// SIMATIC S7-200 project (STEP 7-Micro/WIN), CPU 224XP CN REL 02.01

SYMBOL_TABLE USUARIO1
SO               I0.3     // Sensor de Objetos (Detecta la pieza para iniciar la seleccion)
S_I              I0.4     // Sensor de fibra Optica (clasificacion de materiales)
SM               I0.5     // Sensor magnetico (clasificacion de materiales)
S1               I0.7     // Sensor de retorno del cilindro 1
S2               I1.0     // Sensor de retorno del cilindro 2
S3               I1.1     // Sensor de retorno del cilindro 3
SBB1             I1.3     // Pulsador de Marcha
SBB2             I1.2     // Pulsador de Paro
QS               I1.4     // Zeta de emergencia
SA               I1.5     // Selector rotatorio
am               Q0.0     // Motor
C_1              Q0.4     // cilindro neumatico 1
C_2              Q0.5     // cilindro neumatico 2
C_3              Q0.6     // cilindro neumatico 3
HL1              Q0.7     // Lampara de señalizacion amarilla
HL2              Q1.0     // Lampara de señalizacion verde
HL3              Q1.1     // Lampara de señalizacion roja
E0               M0.0     // Estado 0
E1               M0.1     // Estado 1
E2               M0.2     // Estado 2
E3               M0.3     // Estado 3
E4               M0.4     // Estado 4
E5               M0.5     // Estado 5
E6               M0.6     // Estado 6
E7               M0.7     // Estado 7
E8               M1.0     // Estado 8
E9               M1.1     // Estado 9
E10              M1.2     // Estado 10
E11              M1.3     // Estado 11
E12              M1.4     // Estado 12
E13              M1.5     // Estado 13
E14              M1.6     // Estado 14
EM               M1.7     // Variable para paro momentaneo
MOTOR            M2.0     // Variable para activacion o desactivacion del motor
E15              M2.1     // Estado 15
E16              M2.2     // Estado 16
C_C0             VD110
C_C1             VD100
r_k              VD190
m_k              VD120
m_k_1            VD130
m_k_2            VD140
e_k              VD150
e_k_1            VD160
e_k_2            VD170
Ao               VD200
Bo               VD210
Co               VD220
Do               VD230
Eo               VD240
L_k              VD180
set_point        VD90
END_SYMBOL_TABLE

ORGANIZATION_BLOCK PRINCIPAL:OB1
TITLE=UNIDAD DE SELECCION
BEGIN
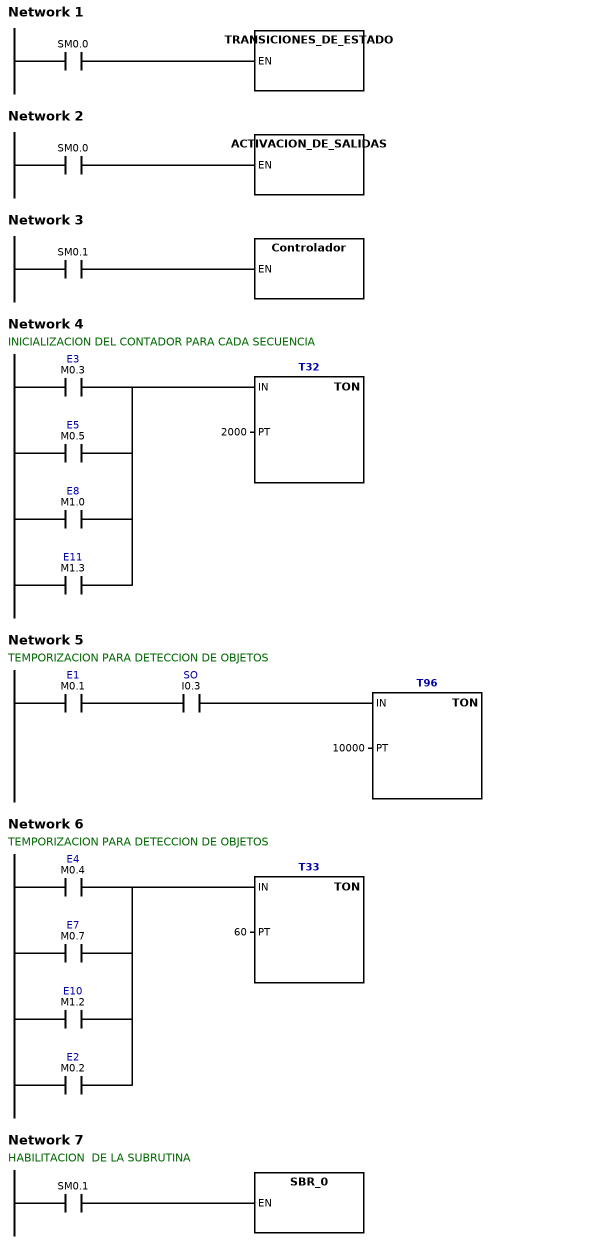
Network 1
LD     SM0.0
CALL   TRANSICIONES_DE_ESTADO:SBR1
Network 2
LD     SM0.0
CALL   ACTIVACION_DE_SALIDAS:SBR2
Network 3
LD     SM0.1
CALL   Controlador:SBR3
Network 4
// INICIALIZACION DEL CONTADOR PARA CADA SECUENCIA 
LD     E3:M0.3
O      E5:M0.5
O      E8:M1.0
O      E11:M1.3
TON    T32, 2000
Network 5
// TEMPORIZACION PARA DETECCION DE OBJETOS
LD     E1:M0.1
A      SO:I0.3
TON    T96, 10000
Network 6
// TEMPORIZACION PARA DETECCION DE OBJETOS
LD     E4:M0.4
O      E7:M0.7
O      E10:M1.2
O      E2:M0.2
TON    T33, 60
Network 7
// HABILITACION  DE LA SUBRUTINA
LD     SM0.1
CALL   SBR_0:SBR0
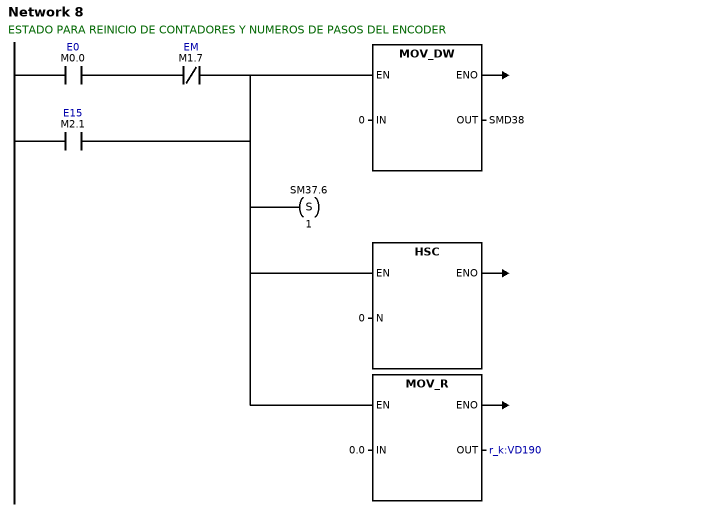
Network 8
// ESTADO PARA REINICIO DE CONTADORES Y NUMEROS DE PASOS DEL ENCODER
LD     E0:M0.0
AN     EM:M1.7
O      E15:M2.1
MOVD   0, SMD38
S      SM37.6, 1
HSC    0
MOVR   0.0, r_k:VD190
END_ORGANIZATION_BLOCK

SUBROUTINE_BLOCK SBR_0:SBR0
TITLE=COMENTARIOS DE LA SUBRUTINA
BEGIN
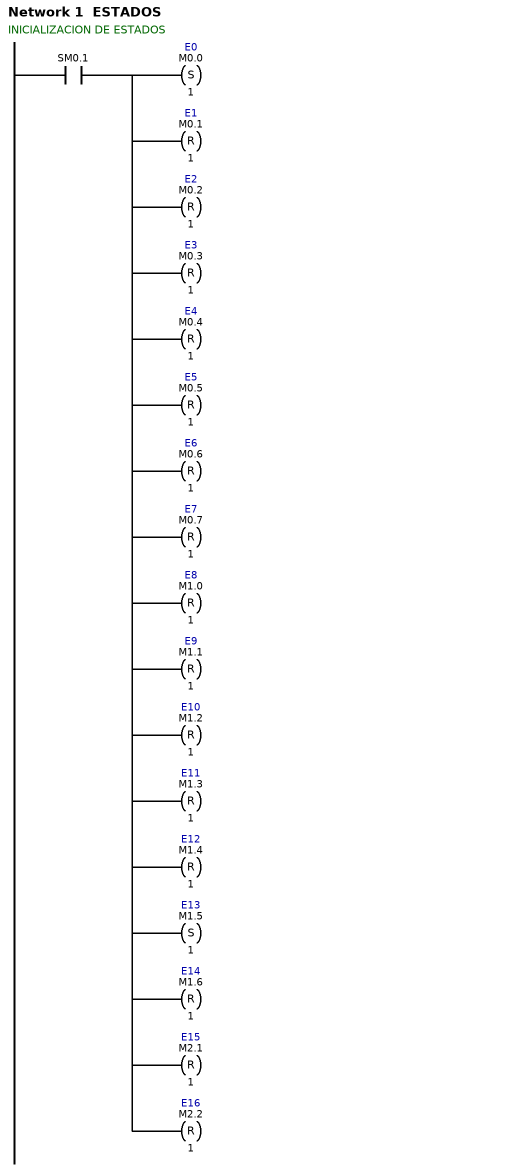
Network 1 // ESTADOS
// INICIALIZACION DE ESTADOS
LD     SM0.1
S      E0:M0.0, 1
R      E1:M0.1, 1
R      E2:M0.2, 1
R      E3:M0.3, 1
R      E4:M0.4, 1
R      E5:M0.5, 1
R      E6:M0.6, 1
R      E7:M0.7, 1
R      E8:M1.0, 1
R      E9:M1.1, 1
R      E10:M1.2, 1
R      E11:M1.3, 1
R      E12:M1.4, 1
S      E13:M1.5, 1
R      E14:M1.6, 1
R      E15:M2.1, 1
R      E16:M2.2, 1
END_SUBROUTINE_BLOCK

SUBROUTINE_BLOCK TRANSICIONES_DE_ESTADO:SBR1
TITLE=TRANSICIONES DE ESTADO
BEGIN
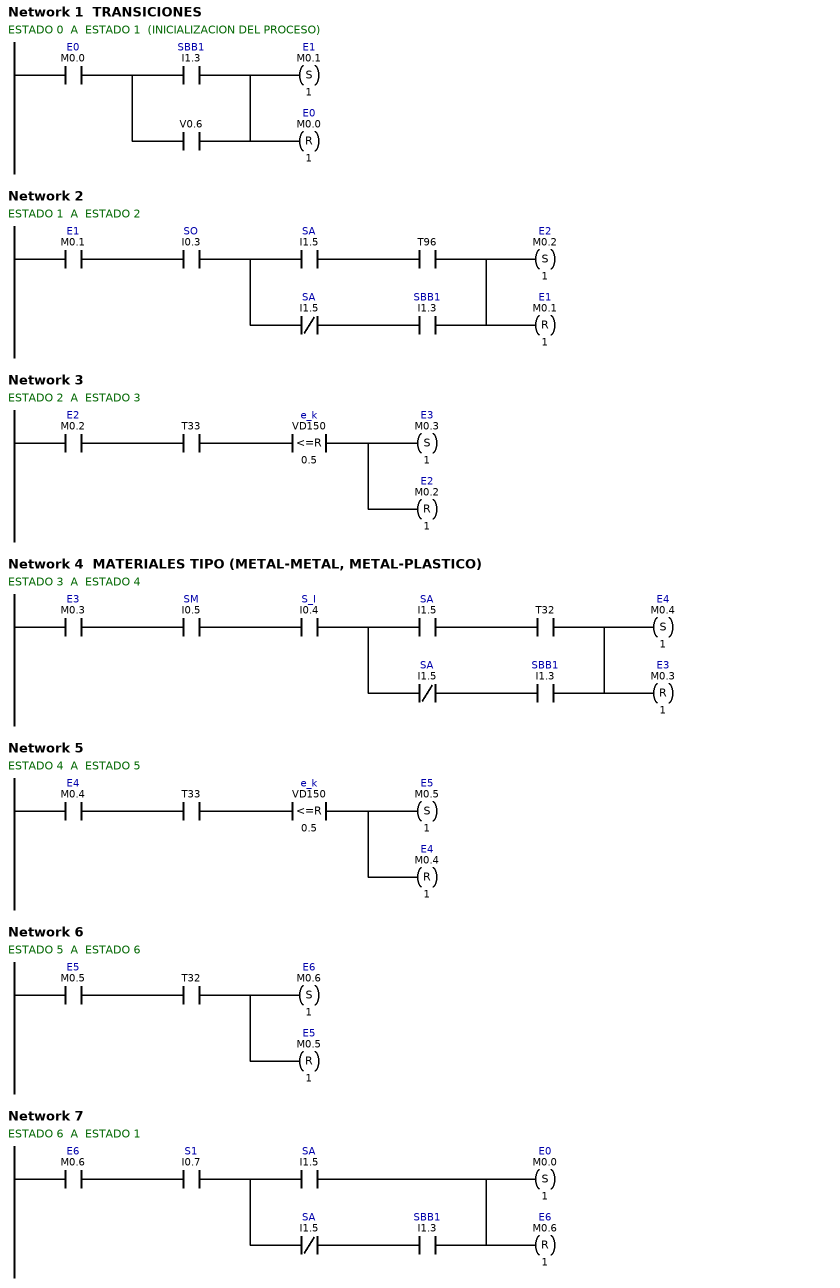
Network 1 // TRANSICIONES
// ESTADO 0  A  ESTADO 1  (INICIALIZACION DEL PROCESO)
LD     E0:M0.0
LD     SBB1:I1.3
O      V0.6
ALD
S      E1:M0.1, 1
R      E0:M0.0, 1
Network 2
// ESTADO 1  A  ESTADO 2 
LD     E1:M0.1
A      SO:I0.3
LD     SA:I1.5
A      T96
LDN    SA:I1.5
A      SBB1:I1.3
OLD
ALD
S      E2:M0.2, 1
R      E1:M0.1, 1
Network 3
// ESTADO 2  A  ESTADO 3
LD     E2:M0.2
A      T33
AR<=   e_k:VD150, 0.5
S      E3:M0.3, 1
R      E2:M0.2, 1
Network 4 // MATERIALES TIPO (METAL-METAL, METAL-PLASTICO)
// ESTADO 3  A  ESTADO 4
LD     E3:M0.3
A      SM:I0.5
A      S_I:I0.4
LD     SA:I1.5
A      T32
LDN    SA:I1.5
A      SBB1:I1.3
OLD
ALD
S      E4:M0.4, 1
R      E3:M0.3, 1
Network 5
// ESTADO 4  A  ESTADO 5
LD     E4:M0.4
A      T33
AR<=   e_k:VD150, 0.5
S      E5:M0.5, 1
R      E4:M0.4, 1
Network 6
// ESTADO 5  A  ESTADO 6
LD     E5:M0.5
A      T32
S      E6:M0.6, 1
R      E5:M0.5, 1
Network 7
// ESTADO 6  A  ESTADO 1
LD     E6:M0.6
A      S1:I0.7
LD     SA:I1.5
LDN    SA:I1.5
A      SBB1:I1.3
OLD
ALD
S      E0:M0.0, 1
R      E6:M0.6, 1
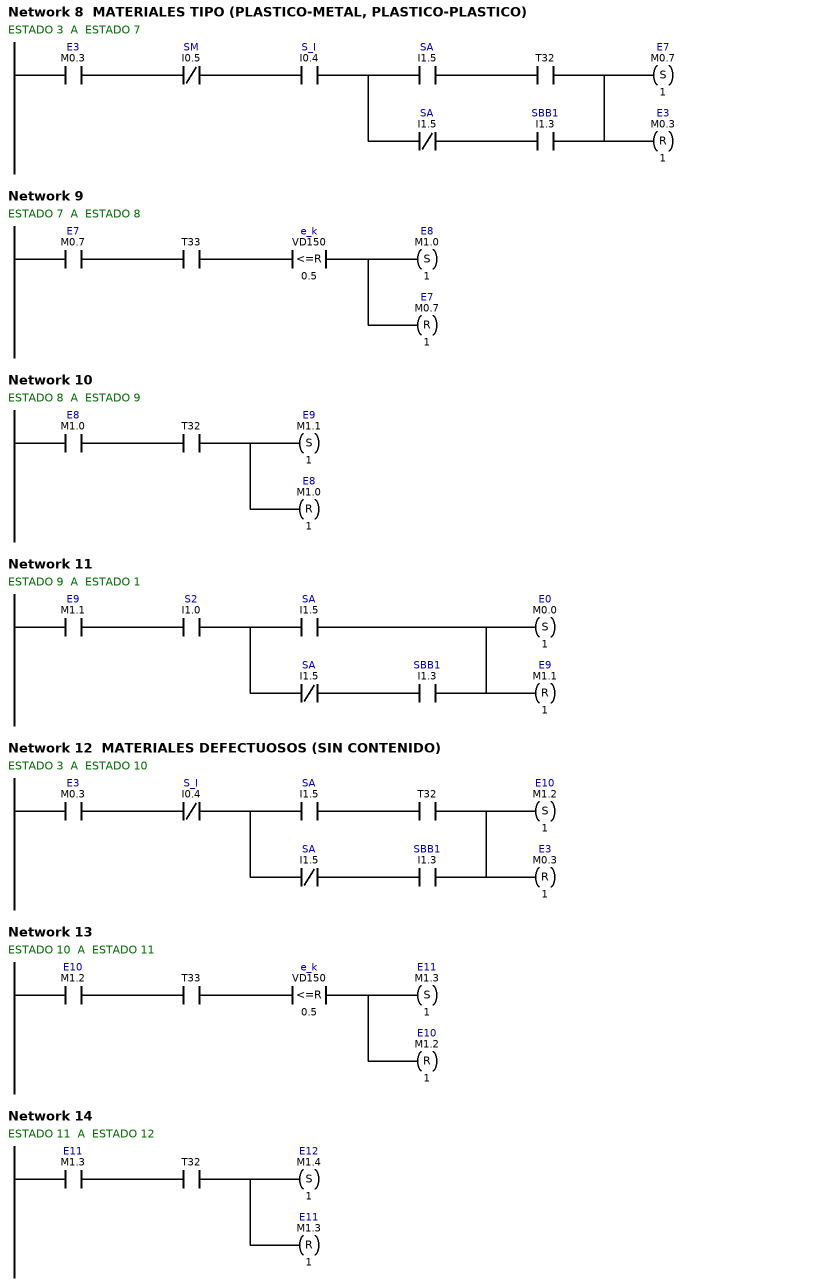
Network 8 // MATERIALES TIPO (PLASTICO-METAL, PLASTICO-PLASTICO)
// ESTADO 3  A  ESTADO 7
LD     E3:M0.3
AN     SM:I0.5
A      S_I:I0.4
LD     SA:I1.5
A      T32
LDN    SA:I1.5
A      SBB1:I1.3
OLD
ALD
S      E7:M0.7, 1
R      E3:M0.3, 1
Network 9
// ESTADO 7  A  ESTADO 8
LD     E7:M0.7
A      T33
AR<=   e_k:VD150, 0.5
S      E8:M1.0, 1
R      E7:M0.7, 1
Network 10
// ESTADO 8  A  ESTADO 9
LD     E8:M1.0
A      T32
S      E9:M1.1, 1
R      E8:M1.0, 1
Network 11
// ESTADO 9  A  ESTADO 1
LD     E9:M1.1
A      S2:I1.0
LD     SA:I1.5
LDN    SA:I1.5
A      SBB1:I1.3
OLD
ALD
S      E0:M0.0, 1
R      E9:M1.1, 1
Network 12 // MATERIALES DEFECTUOSOS (SIN CONTENIDO)
// ESTADO 3  A  ESTADO 10 
LD     E3:M0.3
AN     S_I:I0.4
LD     SA:I1.5
A      T32
LDN    SA:I1.5
A      SBB1:I1.3
OLD
ALD
S      E10:M1.2, 1
R      E3:M0.3, 1
Network 13
// ESTADO 10  A  ESTADO 11
LD     E10:M1.2
A      T33
AR<=   e_k:VD150, 0.5
S      E11:M1.3, 1
R      E10:M1.2, 1
Network 14
// ESTADO 11  A  ESTADO 12
LD     E11:M1.3
A      T32
S      E12:M1.4, 1
R      E11:M1.3, 1
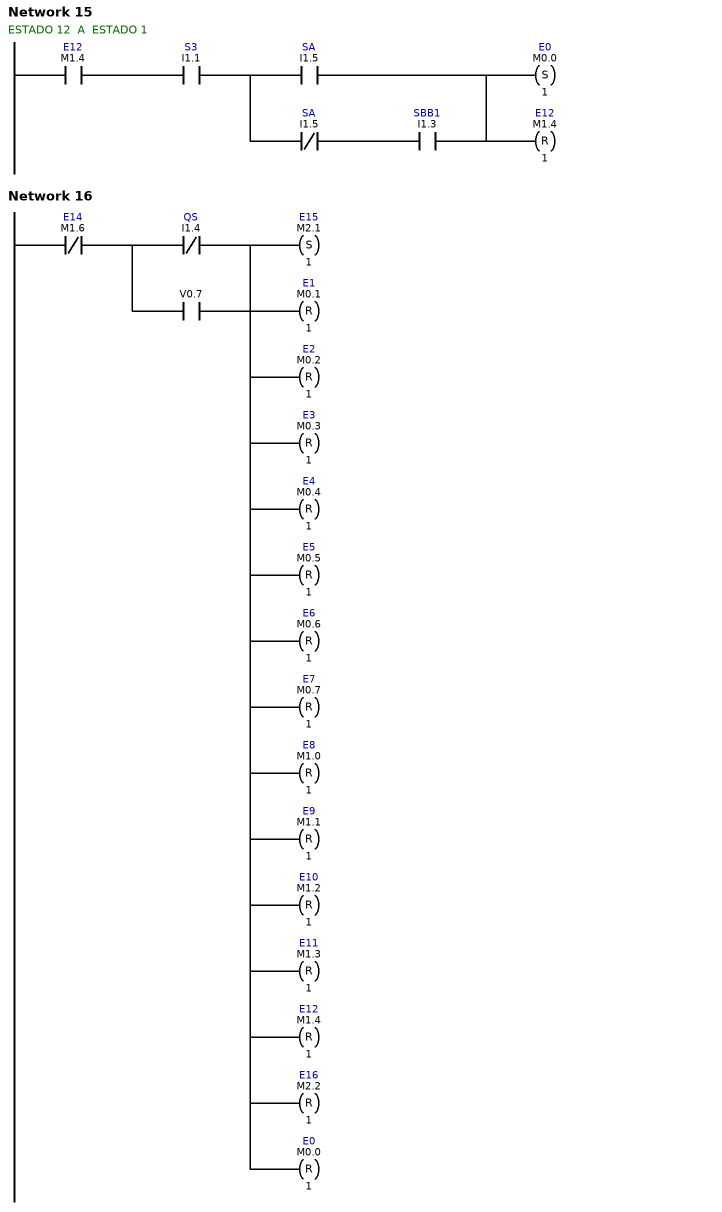
Network 15
// ESTADO 12  A  ESTADO 1
LD     E12:M1.4
A      S3:I1.1
LD     SA:I1.5
LDN    SA:I1.5
A      SBB1:I1.3
OLD
ALD
S      E0:M0.0, 1
R      E12:M1.4, 1
Network 16
LDN    E14:M1.6
LDN    QS:I1.4
O      V0.7
ALD
S      E15:M2.1, 1
R      E1:M0.1, 1
R      E2:M0.2, 1
R      E3:M0.3, 1
R      E4:M0.4, 1
R      E5:M0.5, 1
R      E6:M0.6, 1
R      E7:M0.7, 1
R      E8:M1.0, 1
R      E9:M1.1, 1
R      E10:M1.2, 1
R      E11:M1.3, 1
R      E12:M1.4, 1
R      E16:M2.2, 1
R      E0:M0.0, 1
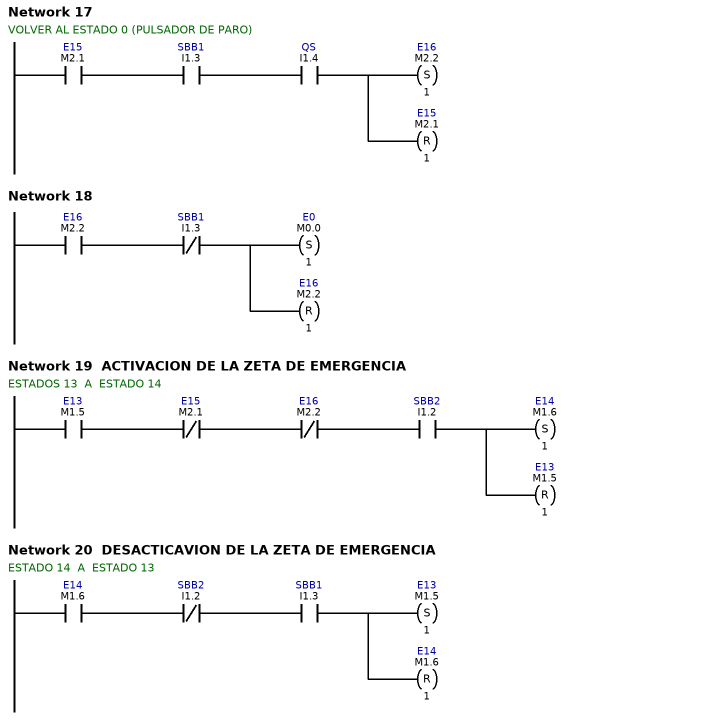
Network 17
// VOLVER AL ESTADO 0 (PULSADOR DE PARO)
LD     E15:M2.1
A      SBB1:I1.3
A      QS:I1.4
S      E16:M2.2, 1
R      E15:M2.1, 1
Network 18
LD     E16:M2.2
AN     SBB1:I1.3
S      E0:M0.0, 1
R      E16:M2.2, 1
Network 19 // ACTIVACION DE LA ZETA DE EMERGENCIA
// ESTADOS 13  A  ESTADO 14
LD     E13:M1.5
AN     E15:M2.1
AN     E16:M2.2
A      SBB2:I1.2
S      E14:M1.6, 1
R      E13:M1.5, 1
Network 20 // DESACTICAVION DE LA ZETA DE EMERGENCIA
// ESTADO 14  A  ESTADO 13
LD     E14:M1.6
AN     SBB2:I1.2
A      SBB1:I1.3
S      E13:M1.5, 1
R      E14:M1.6, 1
Network 21 // Título de segmento
// Comentario de segmento
END_SUBROUTINE_BLOCK

SUBROUTINE_BLOCK ACTIVACION_DE_SALIDAS:SBR2
TITLE=COMENTARIOS DE LA SUBRUTINA
BEGIN
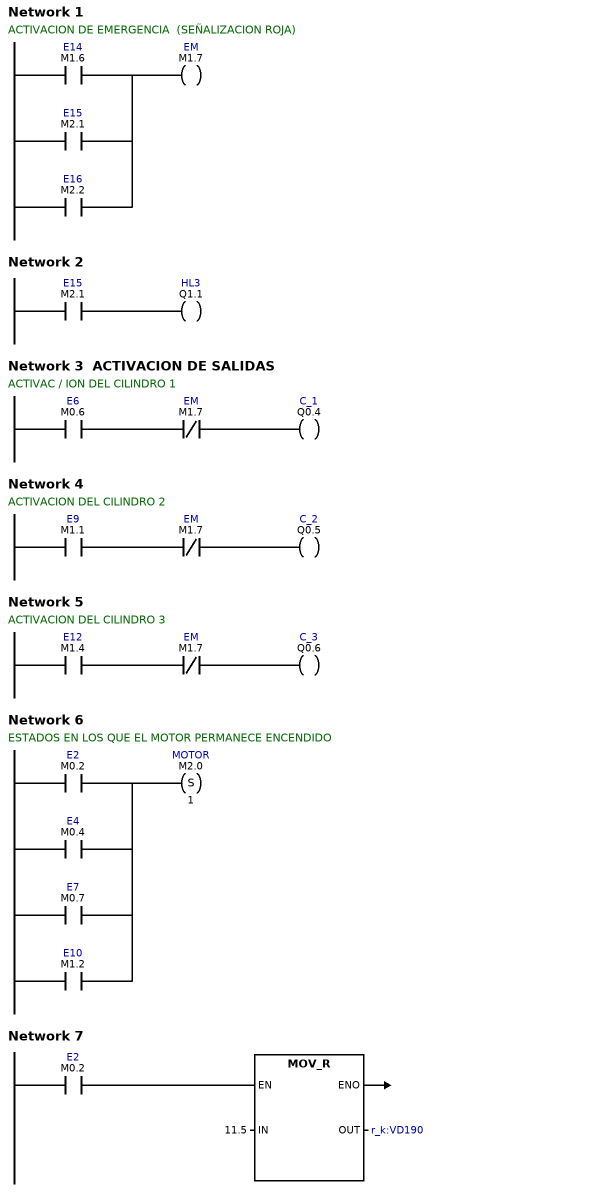
Network 1
// ACTIVACION DE EMERGENCIA  (SEÑALIZACION ROJA)
LD     E14:M1.6
O      E15:M2.1
O      E16:M2.2
=      EM:M1.7
Network 2
LD     E15:M2.1
=      HL3:Q1.1
Network 3 // ACTIVACION DE SALIDAS
// ACTIVAC
// ION DEL CILINDRO 1
LD     E6:M0.6
AN     EM:M1.7
=      C_1:Q0.4
Network 4
// ACTIVACION DEL CILINDRO 2
LD     E9:M1.1
AN     EM:M1.7
=      C_2:Q0.5
Network 5
// ACTIVACION DEL CILINDRO 3
LD     E12:M1.4
AN     EM:M1.7
=      C_3:Q0.6
Network 6
// ESTADOS EN LOS QUE EL MOTOR PERMANECE ENCENDIDO
LD     E2:M0.2
O      E4:M0.4
O      E7:M0.7
O      E10:M1.2
S      MOTOR:M2.0, 1
Network 7
LD     E2:M0.2
MOVR   11.5, r_k:VD190
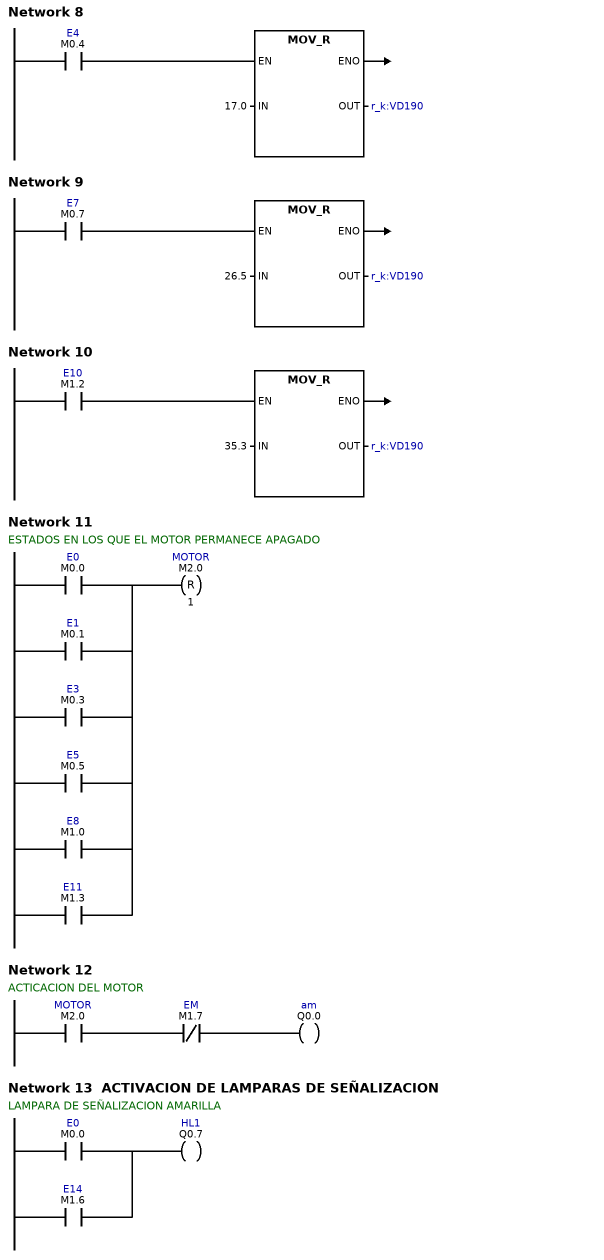
Network 8
LD     E4:M0.4
MOVR   17.0, r_k:VD190
Network 9
LD     E7:M0.7
MOVR   26.5, r_k:VD190
Network 10
LD     E10:M1.2
MOVR   35.3, r_k:VD190
Network 11
// ESTADOS EN LOS QUE EL MOTOR PERMANECE APAGADO
LD     E0:M0.0
O      E1:M0.1
O      E3:M0.3
O      E5:M0.5
O      E8:M1.0
O      E11:M1.3
R      MOTOR:M2.0, 1
Network 12
// ACTICACION DEL MOTOR
LD     MOTOR:M2.0
AN     EM:M1.7
=      am:Q0.0
Network 13 // ACTIVACION DE LAMPARAS DE SEÑALIZACION
// LAMPARA DE SEÑALIZACION AMARILLA
LD     E0:M0.0
O      E14:M1.6
=      HL1:Q0.7
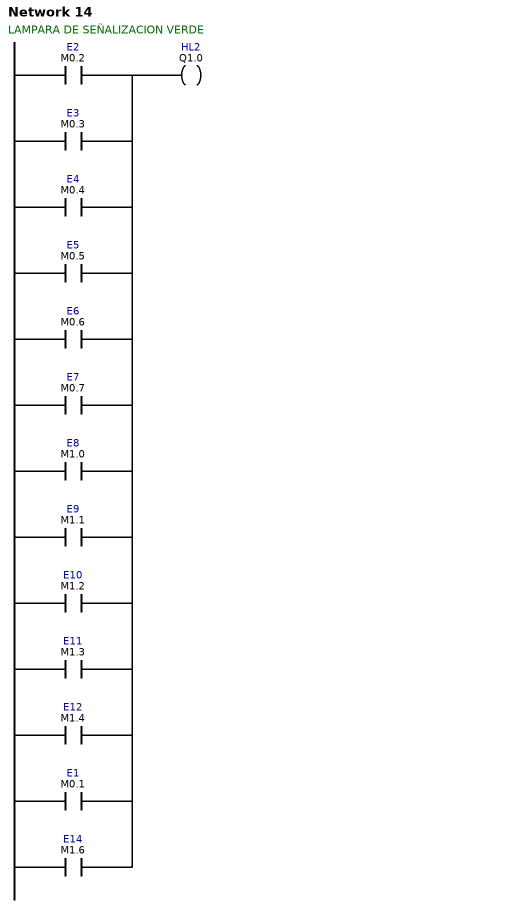
Network 14
// LAMPARA DE SEÑALIZACION VERDE
LD     E2:M0.2
O      E3:M0.3
O      E4:M0.4
O      E5:M0.5
O      E6:M0.6
O      E7:M0.7
O      E8:M1.0
O      E9:M1.1
O      E10:M1.2
O      E11:M1.3
O      E12:M1.4
O      E1:M0.1
O      E14:M1.6
=      HL2:Q1.0
Network 15 // Título de segmento
// Comentario de segmento
END_SUBROUTINE_BLOCK

SUBROUTINE_BLOCK Controlador:SBR3
TITLE=
BEGIN
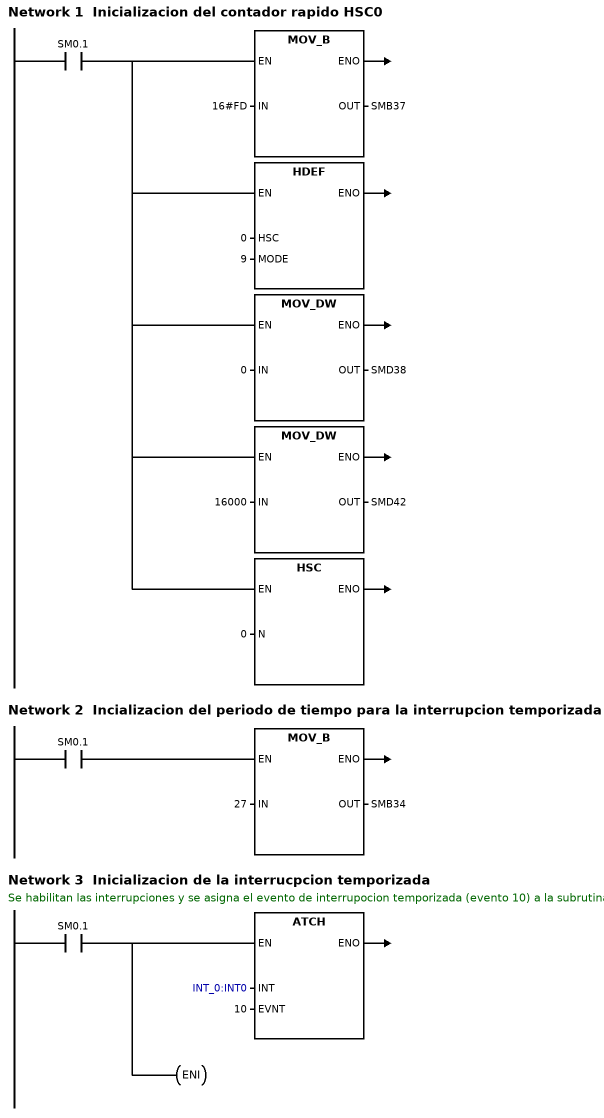
Network 1 // Inicializacion del contador rapido HSC0
LD     SM0.1
MOVB   16#FD, SMB37
HDEF   0, 9
MOVD   0, SMD38
MOVD   16000, SMD42
HSC    0
Network 2 // Incializacion del periodo de tiempo para la interrupcion temporizada
LD     SM0.1
MOVB   27, SMB34
Network 3 // Inicializacion de la interrucpcion temporizada
// Se habilitan las interrupciones y se asigna el evento de interrupocion temporizada (evento 10) a la subrutina de interrupcion INT_0
LD     SM0.1
ATCH   INT_0:INT0, 10
ENI
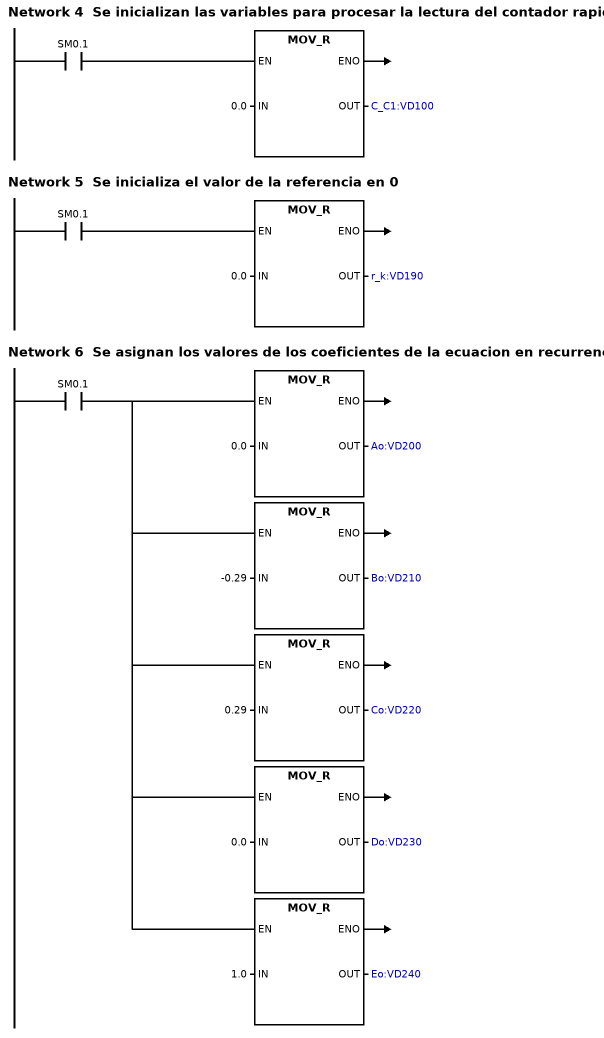
Network 4 // Se inicializan las variables para procesar la lectura del contador rapido HSC0
LD     SM0.1
MOVR   0.0, C_C1:VD100
Network 5 // Se inicializa el valor de la referencia en 0
LD     SM0.1
MOVR   0.0, r_k:VD190
Network 6 // Se asignan los valores de los coeficientes de la ecuacion en recurrencia
LD     SM0.1
MOVR   0.0, Ao:VD200
MOVR   -0.29, Bo:VD210
MOVR   0.29, Co:VD220
MOVR   0.0, Do:VD230
MOVR   1.0, Eo:VD240
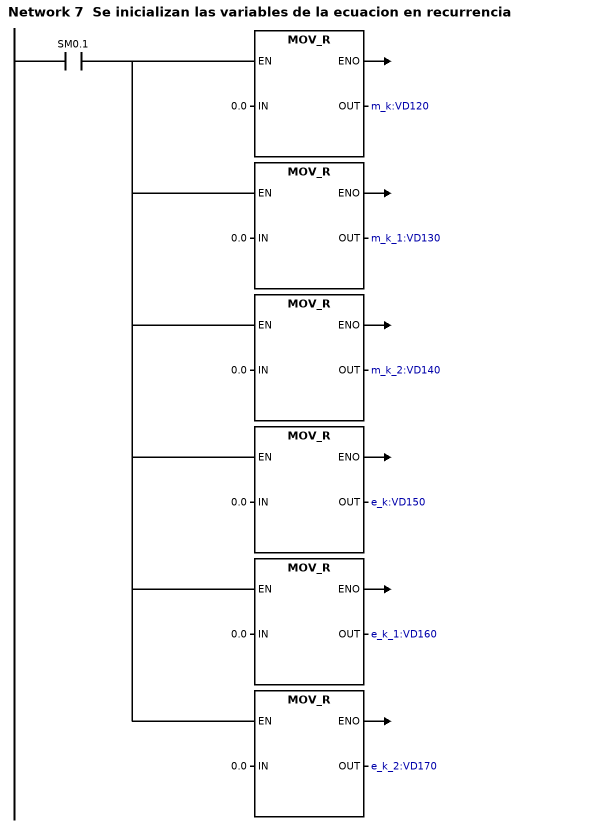
Network 7 // Se inicializan las variables de la ecuacion en recurrencia
LD     SM0.1
MOVR   0.0, m_k:VD120
MOVR   0.0, m_k_1:VD130
MOVR   0.0, m_k_2:VD140
MOVR   0.0, e_k:VD150
MOVR   0.0, e_k_1:VD160
MOVR   0.0, e_k_2:VD170
END_SUBROUTINE_BLOCK

INTERRUPT_BLOCK INT_0:INT0
TITLE=COMENTARIOS DE LA RUTINA DE INTERRUPCIÓN
BEGIN
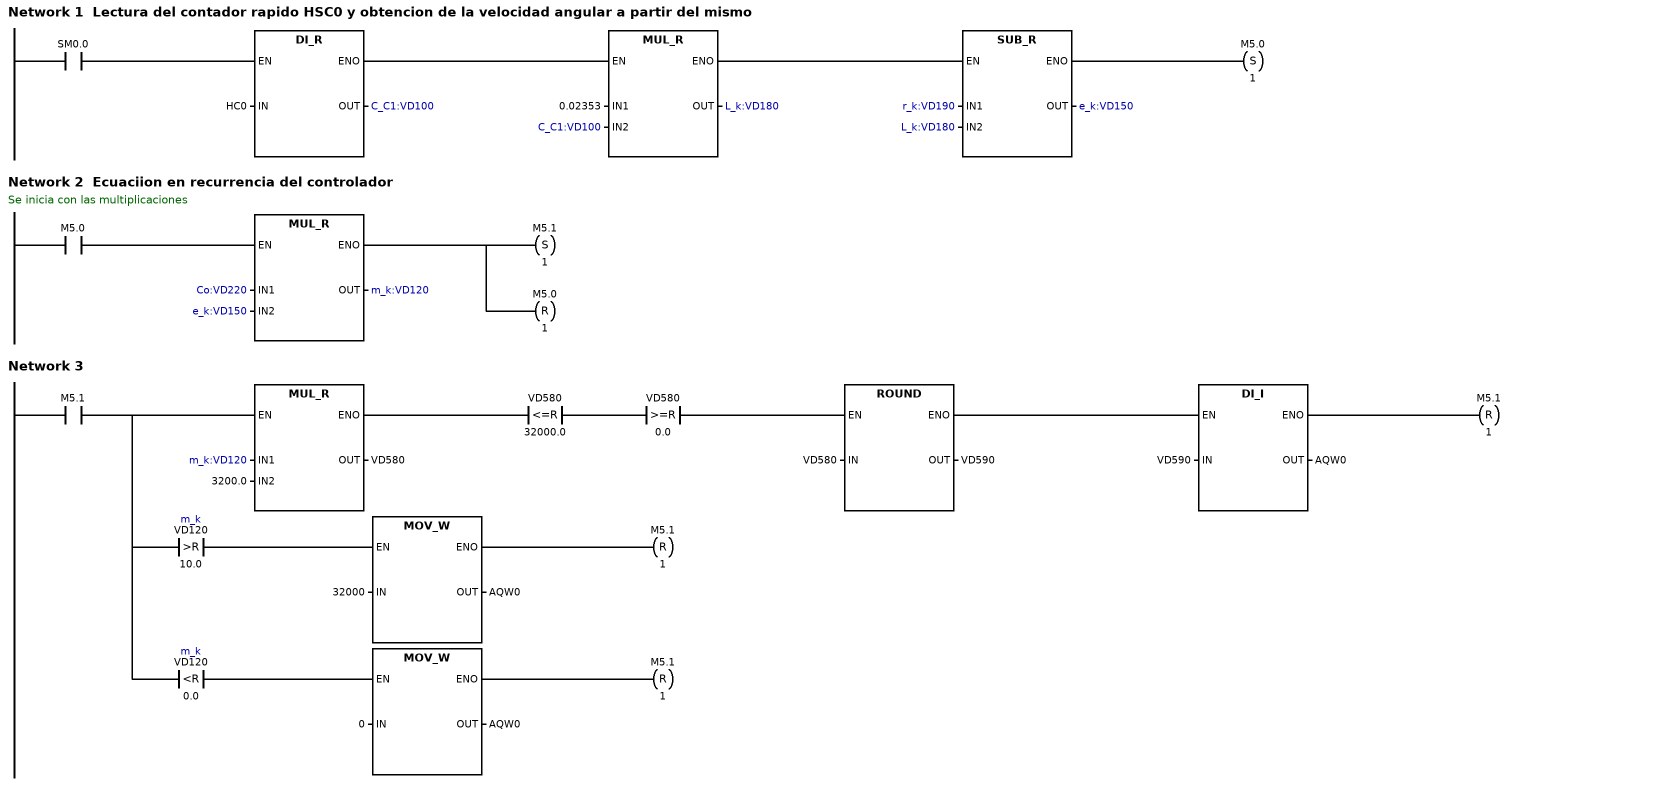
Network 1 // Lectura del contador rapido HSC0 y obtencion de la velocidad angular a partir del mismo
LD     SM0.0
DTR    HC0, C_C1:VD100
AENO
MOVR   0.02353, L_k:VD180
AENO
*R     C_C1:VD100, L_k:VD180
AENO
MOVR   r_k:VD190, e_k:VD150
AENO
-R     L_k:VD180, e_k:VD150
AENO
S      M5.0, 1
Network 2 // Ecuaciion en recurrencia del controlador 
// Se inicia con las multiplicaciones
LD     M5.0
MOVR   Co:VD220, m_k:VD120
AENO
*R     e_k:VD150, m_k:VD120
AENO
S      M5.1, 1
R      M5.0, 1
Network 3
LD     M5.1
LPS
MOVR   m_k:VD120, VD580
AENO
*R     3200.0, VD580
AENO
AR<=   VD580, 32000.0
AR>=   VD580, 0.0
ROUND  VD580, VD590
AENO
DTI    VD590, AQW0
AENO
R      M5.1, 1
LRD
AR>    m_k:VD120, 10.0
MOVW   32000, AQW0
AENO
R      M5.1, 1
LPP
AR<    m_k:VD120, 0.0
MOVW   0, AQW0
AENO
R      M5.1, 1
Network 4 // Título de segmento
// Comentario de segmento
END_INTERRUPT_BLOCK
